FUNCTION_BLOCK ConveyorStationCtrl (* Basic Function Block Type *)
  (* Standard: 61499-2 *)
  (* Version 0.0, 7/2/2026, Template *)
  PACKAGE Main;
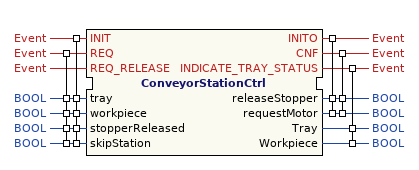
  EVENT_INPUT
    INIT WITH tray, workpiece, stopperReleased, skipStation; (* Initialization Request *)
    REQ WITH tray, workpiece, stopperReleased, skipStation; (* Normal Execution Request *)
    REQ_RELEASE;
  END_EVENT
  EVENT_OUTPUT
    INITO WITH releaseStopper, requestMotor; (* Initialization Confirm *)
    CNF WITH releaseStopper, requestMotor; (* Execution Confirmation *)
    INDICATE_TRAY_STATUS WITH Tray, Workpiece;
  END_EVENT
  VAR_INPUT
    tray : BOOL; (* Input event qualifier *)
    workpiece : BOOL;
    stopperReleased : BOOL;
    skipStation : BOOL;
  END_VAR
  VAR_OUTPUT
    releaseStopper : BOOL; (* Output event qualifier *)
    requestMotor : BOOL;
    Tray : BOOL;
    Workpiece : BOOL;
  END_VAR
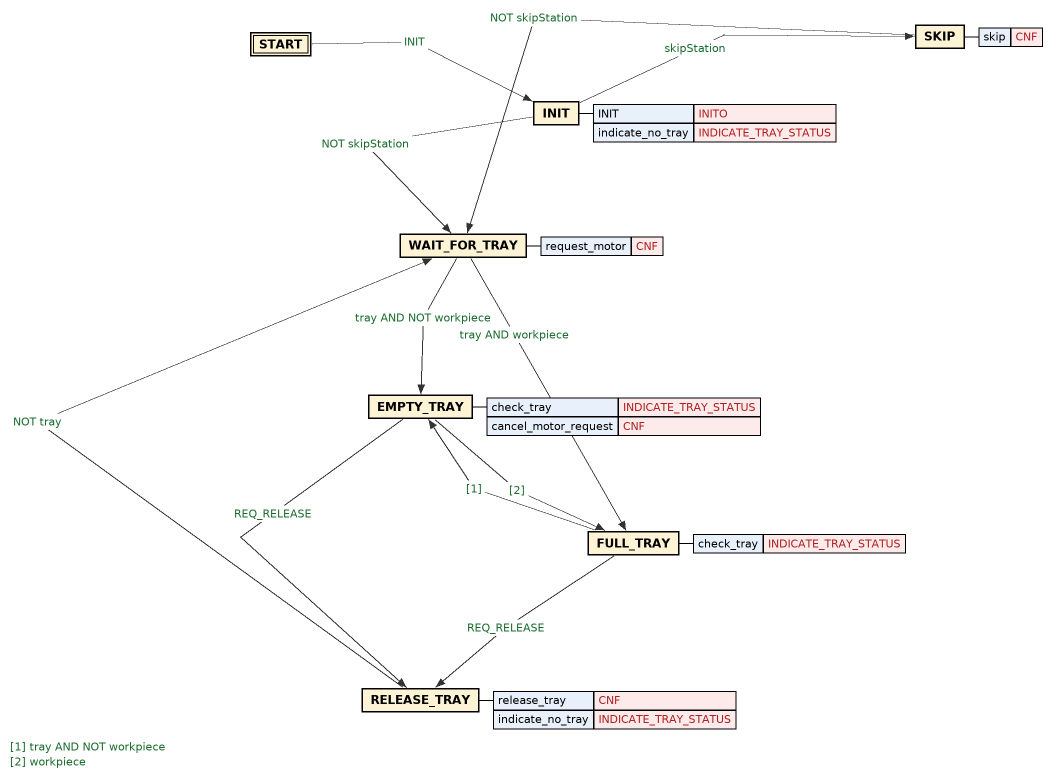
  EC_STATES
    START; (* Initial State *)
    INIT : INIT -> INITO, indicate_no_tray -> INDICATE_TRAY_STATUS; (* Initialization *)
    SKIP : skip -> CNF;
    WAIT_FOR_TRAY : request_motor -> CNF;
    EMPTY_TRAY : check_tray -> INDICATE_TRAY_STATUS, cancel_motor_request -> CNF;
    FULL_TRAY : check_tray -> INDICATE_TRAY_STATUS;
    RELEASE_TRAY : release_tray -> CNF, indicate_no_tray -> INDICATE_TRAY_STATUS;
  END_STATES
  EC_TRANSITIONS
    START TO INIT := INIT;
    INIT TO SKIP := skipStation;
    SKIP TO WAIT_FOR_TRAY := NOT skipStation;
    INIT TO WAIT_FOR_TRAY := NOT skipStation;
    WAIT_FOR_TRAY TO FULL_TRAY := tray AND workpiece;
    WAIT_FOR_TRAY TO EMPTY_TRAY := tray AND NOT workpiece;
    EMPTY_TRAY TO FULL_TRAY := workpiece;
    FULL_TRAY TO EMPTY_TRAY := tray AND NOT workpiece;
    FULL_TRAY TO RELEASE_TRAY := REQ_RELEASE;
    RELEASE_TRAY TO WAIT_FOR_TRAY := NOT tray;
    EMPTY_TRAY TO RELEASE_TRAY := REQ_RELEASE;
  END_TRANSITIONS
  ALGORITHM INIT IN ST: (* Initialization algorithm *)
requestMotor := FALSE;
releaseStopper := FALSE;
Tray := FALSE;
Workpiece := FALSE;
  END_ALGORITHM
  ALGORITHM REQ IN ST: (* Normally executed algorithm *)
;
  END_ALGORITHM
  ALGORITHM skip IN ST:
releaseStopper := TRUE;
  END_ALGORITHM
  ALGORITHM indicate_no_tray IN ST:
Tray := FALSE;
Workpiece := FALSE;
  END_ALGORITHM
  ALGORITHM request_motor IN ST:
requestMotor := TRUE;
releaseStopper := FALSE;
  END_ALGORITHM
  ALGORITHM check_tray IN ST:
Tray := tray;
Workpiece := workpiece;
  END_ALGORITHM
  ALGORITHM cancel_motor_request IN ST:
requestMotor := FALSE;
  END_ALGORITHM
  ALGORITHM release_tray IN ST:
releaseStopper := TRUE;
requestMotor := TRUE;
  END_ALGORITHM
END_FUNCTION_BLOCK
